TYPE ST_EL3312CoeWriteData :
STRUCT
	wIdx: WORD;
	bySubIdx: BYTE;
	bWriteOK: BOOL;
	dwData: DWORD;
	nSize: UDINT;
END_STRUCT
END_TYPE

(* stored: Version 1.1.0.1, ProductVersion 3.1.4024.15
   DUT ST_EL3312CoeWriteData: Id {ca3baa5e-e63d-42eb-80d2-e094c9dc213b} *)
